// TIA Portal project "LAB05" (V16)

(* hardware
DEVICE "S7300/ET200M station_1"  S7-300 station
   slot 0: "Rail_0"  Rail  6ES7 390-1***0-0AA0
   slot 2: "PLC_1"  CPU 313C-2 DP  6ES7 313-6CF03-0AB0  V2.6
      slot 0: "MPI interface_1"  X1
      slot 1: "DP interface_1"  X2
      slot 2: "DI 16/DO 16_1"  DI16/DO16
      slot 4: "Count_1"  Counter
*)

// ===== PLC "PLC_1"  CPU 313C-2 DP =====

VAR_GLOBAL   // PLC tag table "Default tag table"
   "Tag_1" AT %MD14 : DWord;
   "Tag_2" AT %MW12 : Word;
   "Tag_3" AT %MW20 : Word;
END_VAR

DATA_BLOCK "DB100"   // DB100
{ S7_Optimized_Access := 'FALSE' }
VERSION : 0.1
   VAR
      Static_1 : Byte := 16#0;
      Static_2 : Byte;
      Static_3 : Byte;
      Static_4 : Byte;
      Static_5 : Byte;
      Static_6 : Byte;
      Static_7 : Byte;
      Static_8 : Byte;
      Static_9 : Byte;
      Static_10 : Byte;
      Static_11 : Byte;
      Static_12 : Byte;
   END_VAR
BEGIN
END_DATA_BLOCK

FUNCTION "FC7" : Void   // FC7, STL
{ S7_Optimized_Access := 'FALSE' }
VERSION : 0.1
BEGIN

REGION Network 1
         OPN   "DB100";  // open DB100
         L     P#0.0;  // initialize pointer
         T     "Tag_1";  // MD14 is the pointer
         L     DBLG;  // load length of the current DB
         T     "Tag_3";
   AZZE: T     "Tag_2";
         L     0;  // load 0
         T     DBB ["Tag_1"];  // transfer in DBB pointed by MD0
         L     P#1.0;  // increment pointer by 1
         L     "Tag_1";
         +D;
         T     "Tag_1";
         L     "Tag_2";  // load db length
         LOOP  AZZE;  // LOOP decreases by 1 the content of ACCU1 and compares it with 0.
   // If different, the code jumps to the label AZZE
END_REGION
END_FUNCTION

FUNCTION "FC72" : Void   // FC72, STL
{ S7_Optimized_Access := 'FALSE' }
VERSION : 0.1
BEGIN

REGION Network 1
         OPN   "DB100";  // open DB100
         L     P#0.0;  // initialize pointer
         T     "Tag_1";  // MD14 is the pointer
         L     DBLG;  // load length of the current DB
         L     10#2;
         /D;  // divide DBLG by 2 (we're using words not bytes)
         T     "Tag_3";
   AZZE: T     "Tag_2";
         L     0;  // load 0
         T     DBW [ "Tag_1"];  // transfer in DBB pointed by MD0
         L     P#2.0;  // increment pointer by 2, avoiding word overlapping
         L     "Tag_1";
         +D;
         T     "Tag_1";
         L     "Tag_2";  // load db length
         LOOP  AZZE;  // LOOP decreases by 1 the content of ACCU1 and compares it with 0.
   // If different, the code jumps to the label AZZE
END_REGION
END_FUNCTION

FUNCTION "FC73" : Void   // FC73, STL
{ S7_Optimized_Access := 'FALSE' }
VERSION : 0.1
BEGIN

REGION Network 1
         OPN   "DB100";  // open DB100
         L     P#0.0;  // initialize pointer
         T     "Tag_1";  // MD14 is the pointer
         L     DBLG;  // load length of the current DB
         L     10#4;
         /D;  // divide DBLG by 4 (we're using double words not bytes)
         T     "Tag_3";
   AZZE: T     "Tag_2";
         L     0;  // load 0
         T     DBD [ "Tag_1"];  // transfer in DBB pointed by MD0
         L     P#4.0;  // increment pointer by 2, avoiding word overlapping
         L     "Tag_1";
         +D;
         T     "Tag_1";
         L     "Tag_2";  // load db length
         LOOP  AZZE;  // LOOP decreases by 1 the content of ACCU1 and compares it with 0.
   // If different, the code jumps to the label AZZE
END_REGION
END_FUNCTION

ORGANIZATION_BLOCK "Main"   // OB1, STL
TITLE = "Main Program Sweep (Cycle)"
{ S7_Optimized_Access := 'FALSE' }
VERSION : 0.1
   VAR_TEMP
      OB1_EV_CLASS : Byte;   // Bits 0-3 = 1 (Coming event), Bits 4-7 = 1 (Event class 1)
      OB1_SCAN_1 : Byte;   // 1 (Cold restart scan 1 of OB 1), 3 (Scan 2-n of OB 1)
      OB1_PRIORITY : Byte;   // Priority of OB Execution
      OB1_OB_NUMBR : Byte;   // 1 (Organization block 1, OB1)
      OB1_RESERVED_1 : Byte;   // Reserved for system
      OB1_RESERVED_2 : Byte;   // Reserved for system
      OB1_PREV_CYCLE : Int;   // Cycle time of previous OB1 scan (milliseconds)
      OB1_MIN_CYCLE : Int;   // Minimum cycle time of OB1 (milliseconds)
      OB1_MAX_CYCLE : Int;   // Maximum cycle time of OB1 (milliseconds)
      OB1_DATE_TIME : Date_And_Time;   // Date and time OB1 started
   END_VAR
BEGIN

REGION Network 1
         CALL  "FC73";
END_REGION
END_ORGANIZATION_BLOCK